FUNCTION "fc_chamadasBancos_BT2" : Void
TITLE = fc_chamadasBancos_BT2 v0.1
{ S7_Optimized_Access := 'TRUE' }
AUTHOR : 'Reginaldo Lobo'
VERSION : 0.1
////====================================
//// fc_chamadasBancos_BT2 v0.1 (03/11/2026) - GERADO por gerar_banco_v0.2.py - RASCUNHO, nao compilado
//// ONDE RODA : 1515 (BT2). Chamar 1x por ciclo no OB1: "fc_chamadasBancos_BT2"();   (substitui colar chamadas uma a uma)
//// O QUE FAZ : para cada banco, 1) comunicacao com o ET200 (FB101/FB103) e 2) setup das chaves (FB100/FB102), nessa ordem.
//// OBS       : todos os bancos usam a MESMA conexao S7 (W#16#100), decisao do operador de 03/11/2026.
//// ATENCAO   : os DBs de instancia (db30x4i_.../db30x5i_...) precisam existir com esses nomes (criar no TIA como instancia dos FBs).
////=====================================
BEGIN

   // ---------------- BC56 (13 chaves, FB100/101) ----------------
   "db3005i_BC56_ComEt200"(Hab := TRUE, ID_Conexao := W#16#100,
       RemotoCmd := P#DB38.DBX0.0 BYTE 6, RemotoFb := P#DB38.DBX6.0 BYTE 6,
       ComOk => "db3000_BC56_Chaves".sbBanco.comEt200Ok, SeletoraAuto => "db3000_BC56_Chaves".sbBanco.seletoraAuto,
       CbLigar := "db3000_BC56_Chaves".cb.ligar, SbLigada := "db3000_BC56_Chaves".sb.ligada, LigarBanco := "db3000_BC56_Chaves".cbBanco.ligar);

   "db3004i_BC56_SetupChaves"(
       NumChaves := 13, GeradorOperando := "db52_BancoTeste2_DSE".ledManual, EnsaioAtivo := FALSE,   // TODO: tag real do DB "Dados do ensaio"
       kWMedido := "db52_BancoTeste2_DSE".potenciaKw, VaMedido := "db52_BancoTeste2_DSE".tensaoL1L2,
       VbMedido := "db52_BancoTeste2_DSE".tensaoL2L3, VcMedido := "db52_BancoTeste2_DSE".tensaoL3L1,
       TensaoSel := "db3002_BC56_SetupPorTensao".selV.tensaoSel, ChaveSelecionada := "db3000_BC56_Chaves".setup.chaveSel, ComandoSalvar := "db3000_BC56_Chaves".setup.salvar,
       kWNominal := "db3000_BC56_Chaves".setup.nominal, CbLigar := "db3000_BC56_Chaves".cb.ligar, SbLigada := "db3000_BC56_Chaves".sb.ligada, Habilitada := "db3000_BC56_Chaves".setup.habilitada,
       SetupOk := "db3000_BC56_Chaves".setup.setupOk, KwReal := "db3000_BC56_Chaves".setup.kwReal, RmedidoOhm := "db3000_BC56_Chaves".setup.rMedidoOhm,
       RteoricoOhm := "db3000_BC56_Chaves".setup.rTeoricoOhm, SetupData := "db3000_BC56_Chaves".setup.setupData,
       KwRealV := "db3002_BC56_SetupPorTensao".setupV.kwReal, RmedidoV := "db3002_BC56_SetupPorTensao".setupV.rMedidoOhm, VmedidaV := "db3002_BC56_SetupPorTensao".setupV.vMedidaV,
       BaseKwV := "db3002_BC56_SetupPorTensao".setupV.baseKw, SetupDataV := "db3002_BC56_SetupPorTensao".setupV.setupData, SetupOkV := "db3002_BC56_SetupPorTensao".setupV.setupOk);

   // ---------------- BC400 (13 chaves, FB100/101) ----------------
   "db3105i_BC400_ComEt200"(Hab := TRUE, ID_Conexao := W#16#100,
       RemotoCmd := P#DB39.DBX0.0 BYTE 6, RemotoFb := P#DB39.DBX6.0 BYTE 6,
       ComOk => "db3100_BC400_Chaves".sbBanco.comEt200Ok, SeletoraAuto => "db3100_BC400_Chaves".sbBanco.seletoraAuto,
       CbLigar := "db3100_BC400_Chaves".cb.ligar, SbLigada := "db3100_BC400_Chaves".sb.ligada, LigarBanco := "db3100_BC400_Chaves".cbBanco.ligar);

   "db3104i_BC400_SetupChaves"(
       NumChaves := 13, GeradorOperando := "db52_BancoTeste2_DSE".ledManual, EnsaioAtivo := FALSE,   // TODO: tag real do DB "Dados do ensaio"
       kWMedido := "db52_BancoTeste2_DSE".potenciaKw, VaMedido := "db52_BancoTeste2_DSE".tensaoL1L2,
       VbMedido := "db52_BancoTeste2_DSE".tensaoL2L3, VcMedido := "db52_BancoTeste2_DSE".tensaoL3L1,
       TensaoSel := "db3102_BC400_SetupPorTensao".selV.tensaoSel, ChaveSelecionada := "db3100_BC400_Chaves".setup.chaveSel, ComandoSalvar := "db3100_BC400_Chaves".setup.salvar,
       kWNominal := "db3100_BC400_Chaves".setup.nominal, CbLigar := "db3100_BC400_Chaves".cb.ligar, SbLigada := "db3100_BC400_Chaves".sb.ligada, Habilitada := "db3100_BC400_Chaves".setup.habilitada,
       SetupOk := "db3100_BC400_Chaves".setup.setupOk, KwReal := "db3100_BC400_Chaves".setup.kwReal, RmedidoOhm := "db3100_BC400_Chaves".setup.rMedidoOhm,
       RteoricoOhm := "db3100_BC400_Chaves".setup.rTeoricoOhm, SetupData := "db3100_BC400_Chaves".setup.setupData,
       KwRealV := "db3102_BC400_SetupPorTensao".setupV.kwReal, RmedidoV := "db3102_BC400_SetupPorTensao".setupV.rMedidoOhm, VmedidaV := "db3102_BC400_SetupPorTensao".setupV.vMedidaV,
       BaseKwV := "db3102_BC400_SetupPorTensao".setupV.baseKw, SetupDataV := "db3102_BC400_SetupPorTensao".setupV.setupData, SetupOkV := "db3102_BC400_SetupPorTensao".setupV.setupOk);

   // ---------------- BC59,5 (18 chaves, FB102/103) ----------------
   "db3205i_BC595_ComEt200"(Hab := TRUE, ID_Conexao := W#16#100,
       RemotoCmd := P#DB40.DBX0.0 BYTE 8, RemotoFb := P#DB40.DBX8.0 BYTE 8,
       ComOk => "db3200_BC595_Chaves".sbBanco.comEt200Ok, SeletoraAuto => "db3200_BC595_Chaves".sbBanco.seletoraAuto,
       CbLigar := "db3200_BC595_Chaves".cb.ligar, SbLigada := "db3200_BC595_Chaves".sb.ligada, LigarBanco := "db3200_BC595_Chaves".cbBanco.ligar);

   "db3204i_BC595_SetupChaves"(
       NumChaves := 18, GeradorOperando := "db52_BancoTeste2_DSE".ledManual, EnsaioAtivo := FALSE,   // TODO: tag real do DB "Dados do ensaio"
       kWMedido := "db52_BancoTeste2_DSE".potenciaKw, VaMedido := "db52_BancoTeste2_DSE".tensaoL1L2,
       VbMedido := "db52_BancoTeste2_DSE".tensaoL2L3, VcMedido := "db52_BancoTeste2_DSE".tensaoL3L1,
       TensaoSel := "db3202_BC595_SetupPorTensao".selV.tensaoSel, ChaveSelecionada := "db3200_BC595_Chaves".setup.chaveSel, ComandoSalvar := "db3200_BC595_Chaves".setup.salvar,
       kWNominal := "db3200_BC595_Chaves".setup.nominal, CbLigar := "db3200_BC595_Chaves".cb.ligar, SbLigada := "db3200_BC595_Chaves".sb.ligada, Habilitada := "db3200_BC595_Chaves".setup.habilitada,
       SetupOk := "db3200_BC595_Chaves".setup.setupOk, KwReal := "db3200_BC595_Chaves".setup.kwReal, RmedidoOhm := "db3200_BC595_Chaves".setup.rMedidoOhm,
       RteoricoOhm := "db3200_BC595_Chaves".setup.rTeoricoOhm, SetupData := "db3200_BC595_Chaves".setup.setupData,
       KwRealV := "db3202_BC595_SetupPorTensao".setupV.kwReal, RmedidoV := "db3202_BC595_SetupPorTensao".setupV.rMedidoOhm, VmedidaV := "db3202_BC595_SetupPorTensao".setupV.vMedidaV,
       BaseKwV := "db3202_BC595_SetupPorTensao".setupV.baseKw, SetupDataV := "db3202_BC595_SetupPorTensao".setupV.setupData, SetupOkV := "db3202_BC595_SetupPorTensao".setupV.setupOk);

   // ---------------- BC550 (12 chaves, FB100/101) ----------------
   "db3305i_BC550_ComEt200"(Hab := TRUE, ID_Conexao := W#16#100,
       RemotoCmd := P#DB41.DBX0.0 BYTE 6, RemotoFb := P#DB41.DBX6.0 BYTE 6,
       ComOk => "db3300_BC550_Chaves".sbBanco.comEt200Ok, SeletoraAuto => "db3300_BC550_Chaves".sbBanco.seletoraAuto,
       CbLigar := "db3300_BC550_Chaves".cb.ligar, SbLigada := "db3300_BC550_Chaves".sb.ligada, LigarBanco := "db3300_BC550_Chaves".cbBanco.ligar);

   "db3304i_BC550_SetupChaves"(
       NumChaves := 12, GeradorOperando := "db52_BancoTeste2_DSE".ledManual, EnsaioAtivo := FALSE,   // TODO: tag real do DB "Dados do ensaio"
       kWMedido := "db52_BancoTeste2_DSE".potenciaKw, VaMedido := "db52_BancoTeste2_DSE".tensaoL1L2,
       VbMedido := "db52_BancoTeste2_DSE".tensaoL2L3, VcMedido := "db52_BancoTeste2_DSE".tensaoL3L1,
       TensaoSel := "db3302_BC550_SetupPorTensao".selV.tensaoSel, ChaveSelecionada := "db3300_BC550_Chaves".setup.chaveSel, ComandoSalvar := "db3300_BC550_Chaves".setup.salvar,
       kWNominal := "db3300_BC550_Chaves".setup.nominal, CbLigar := "db3300_BC550_Chaves".cb.ligar, SbLigada := "db3300_BC550_Chaves".sb.ligada, Habilitada := "db3300_BC550_Chaves".setup.habilitada,
       SetupOk := "db3300_BC550_Chaves".setup.setupOk, KwReal := "db3300_BC550_Chaves".setup.kwReal, RmedidoOhm := "db3300_BC550_Chaves".setup.rMedidoOhm,
       RteoricoOhm := "db3300_BC550_Chaves".setup.rTeoricoOhm, SetupData := "db3300_BC550_Chaves".setup.setupData,
       KwRealV := "db3302_BC550_SetupPorTensao".setupV.kwReal, RmedidoV := "db3302_BC550_SetupPorTensao".setupV.rMedidoOhm, VmedidaV := "db3302_BC550_SetupPorTensao".setupV.vMedidaV,
       BaseKwV := "db3302_BC550_SetupPorTensao".setupV.baseKw, SetupDataV := "db3302_BC550_SetupPorTensao".setupV.setupData, SetupOkV := "db3302_BC550_SetupPorTensao".setupV.setupOk);
END_FUNCTION
